// TIA Portal V20 export
Screen "Tool Stand Bit"  395x650
  ScreenItem "Robot Name" at 2,2 size 393x48  Type=HmiIOField
  ScreenItem "Background" at -1,49 size 395x601  Type=HmiRectangle
  ScreenItem "Cancel Mode" at 315,4 size 76x42  Type=HmiButton
  ScreenItem "矩形_4" at 34,58 size 324x583  Type=HmiRectangle
  ScreenItem "Text Filed E- Stop_17" at 40,321 size 148x21  Type=HmiTextBox
  ScreenItem "Text Field In Auto On_9" at 40,86 size 148x21  Type=HmiTextBox
  ScreenItem "Text Field Home Position_17" at 40,109 size 148x21  Type=HmiTextBox
  ScreenItem "Text field Robot Status_5" at 34,57 size 324x26  Type=HmiTextBox
  ScreenItem "Text Field Manual_17" at 40,251 size 148x21  Type=HmiTextBox
  ScreenItem "Text Field System Ready_9" at 40,133 size 148x21  Type=HmiTextBox
  ScreenItem "Text Field Motor On_9" at 40,156 size 148x21  Type=HmiTextBox
  ScreenItem "Text Field In Cycle_9" at 40,180 size 148x21  Type=HmiTextBox
  ScreenItem "Text Field Cycle On_17" at 40,203 size 148x21  Type=HmiTextBox
  ScreenItem "Text Field On Path_17" at 40,227 size 148x21  Type=HmiTextBox
  ScreenItem "Text Field Tryout Mode_17" at 40,274 size 148x21  Type=HmiTextBox
  ScreenItem "Text Field Stop_17" at 40,298 size 148x21  Type=HmiTextBox
  ScreenItem "Text Filed Error_9" at 40,345 size 148x21  Type=HmiTextBox
  ScreenItem "Text Filed Process Fault_9" at 40,368 size 148x21  Type=HmiTextBox
  ScreenItem "Text Field Home Position_18" at 40,392 size 148x21  Type=HmiTextBox
  ScreenItem "Text Filed E- Stop_18" at 201,109 size 148x21  Type=HmiTextBox
  ScreenItem "Text Field Manual_18" at 40,463 size 148x21  Type=HmiTextBox
  ScreenItem "Text Field Cycle On_18" at 40,416 size 148x21  Type=HmiTextBox
  ScreenItem "Text Field On Path_18" at 40,439 size 148x21  Type=HmiTextBox
  ScreenItem "Text Field Tryout Mode_18" at 40,486 size 148x21  Type=HmiTextBox
  ScreenItem "Text Field Stop_18" at 201,85 size 148x21  Type=HmiTextBox
  ScreenItem "Text Filed E- Stop_19" at 201,273 size 148x21  Type=HmiTextBox
  ScreenItem "Text Field In Auto On_10" at 201,133 size 148x21  Type=HmiTextBox
  ScreenItem "Text Field Home Position_19" at 201,156 size 148x21  Type=HmiTextBox
  ScreenItem "Text Field System Ready_10" at 201,179 size 148x21  Type=HmiTextBox
  ScreenItem "Text Field Motor On_10" at 201,202 size 148x21  Type=HmiTextBox
  ScreenItem "Text Field Tryout Mode_19" at 201,226 size 148x21  Type=HmiTextBox
  ScreenItem "Text Field Stop_19" at 201,248 size 148x21  Type=HmiTextBox
  ScreenItem "Text Filed Error_10" at 201,297 size 148x21  Type=HmiTextBox
  ScreenItem "Text Filed Process Fault_10" at 201,320 size 148x21  Type=HmiTextBox
  ScreenItem "Text Field Home Position_20" at 201,344 size 148x21  Type=HmiTextBox
  ScreenItem "Text Filed E- Stop_20" at 201,486 size 148x21  Type=HmiTextBox
  ScreenItem "Text Field Manual_20" at 201,415 size 148x21  Type=HmiTextBox
  ScreenItem "Text Field Cycle On_20" at 201,368 size 148x21  Type=HmiTextBox
  ScreenItem "Text Field On Path_20" at 201,391 size 148x21  Type=HmiTextBox
  ScreenItem "Text Field Tryout Mode_20" at 201,438 size 148x21  Type=HmiTextBox
  ScreenItem "Text Field Stop_20" at 201,462 size 148x21  Type=HmiTextBox
  ScreenItem "Text field Robot Status_1" at 34,529 size 324x26  Type=HmiTextBox
  ScreenItem "Text Field In Auto On_1" at 40,561 size 148x21  Type=HmiTextBox
  ScreenItem "Text Field Home Position_1" at 40,584 size 148x21  Type=HmiTextBox
  ScreenItem "Text Field System Ready_1" at 40,608 size 148x21  Type=HmiTextBox
  ScreenItem "Text Field In Auto On_2" at 201,561 size 148x21  Type=HmiTextBox
  ScreenItem "Text Field Home Position_2" at 201,584 size 148x21  Type=HmiTextBox
  ScreenItem "Text Field System Ready_2" at 201,608 size 148x21  Type=HmiTextBox
